Fanuc KAREL source: KB00073.KL

PROGRAM KB00073
%NOLOCKGROUP
VAR
  P1: INTEGER
  P2: STRING[80]
BEGIN
  P1 = 1
  P2 = 'A'
  FORCE_LINK(P1, P2)
END KB00073
